// TIA Portal V20 export
// export: Created 2026-10-20T12:43:26.7862005Z, ExportSetting WithDefaults, DisplayName Totally Integrated Automation Portal, DisplayVersion V20 Update 6, DisplayName TIA Portal Openness, DisplayVersion V20 Update 6, DisplayName TIA Portal Version Control Interface, DisplayVersion V20 Update 6, DisplayName SINAMICS Startdrive Advanced, DisplayVersion V20 SP1, DisplayName SINAMICS Startdrive G130, G150, S120, S150, SINAMICS MV, G220, S200, S210, DisplayVersion V20 SP1, DisplayName SINAMICS Startdrive G110M, G120, G120C, G120D, G120P, G115D, DisplayVersion V20 SP1, DisplayName STEP 7 Professional, DisplayVersion V20 Update 6, DisplayName STEP 7 Safety, DisplayVersion V20 Update 2, DisplayName WinCC Basic/Comfort/Advanced, DisplayVersion V20 Update 6, DisplayName WinCC Unified, DisplayVersion V20 Update 6
DATA_BLOCK "C5104_FB_DB"   // DB125
AUTHOR : Mertin Coetzee
VERSION : 0.1
// stored: AutoNumber true, DBAccessibleFromOPCUA true, InstanceOfName Buffer_Conveyor_FB, InstanceOfType FB
"Buffer_Conveyor_FB"
   // VAR_INPUT
   //    Cnv_Settings : "Buffer_Cnv_Settings";
   //    VTD_Level : UInt;
   //    Safety_OK_Delayed : Bool;
   //    Safety_OK : Bool;
   //    CNV_In_Out : Bool;
   //    LGX_ReadyToSend : Bool;
   //    LGX_ReadyToReceive : Bool;
   // END_VAR
   // VAR_IN_OUT
   //    Cnv_Control : "Buffer_Cnv_Control";
   //    SinaSpeed : SinaSpeed;
   // END_VAR
   // VAR
   //    State : UInt;
   //    Timer_Transfer { S7_SetPoint := 'True'} : TON_TIME;
   //    Watchdog { S7_SetPoint := 'True'} : TON_TIME;
   //    Transfer_Direction { S7_SetPoint := 'True'} : String;
   //    MainSetpoint : Int;
   //    T_Outbound_DB { S7_SetPoint := 'True'} : TON_TIME;
   //    R_TRIG_Instance { S7_SetPoint := 'True'} : R_TRIG;
   //    R_Start_DB { S7_SetPoint := 'True'} : R_TRIG;
   //    R_Stop_DB { S7_SetPoint := 'True'} : R_TRIG;
   //    ID_Decoded { S7_SetPoint := 'True'} : "ID_Decoded";
   //    ID_Decoded_From { S7_SetPoint := 'True'} : "ID_Decoded";
   //    ID_Decoded_To { S7_SetPoint := 'True'} : "ID_Decoded";
   //    R_Slow { S7_SetPoint := 'True'} : R_TRIG;
   //    T_Ramp { S7_SetPoint := 'True'} : TON_TIME;
   //    T_Ramp_In : Bool;
   //    HMI_Reset : Bool;
   //    TCheck_PalletType { S7_SetPoint := 'True'} : TON_TIME;
   // END_VAR
BEGIN
END_DATA_BLOCK
